INTERFACE ITF_Buffer2_4

METHOD Aborted : BOOL
VAR_INPUT
END_VAR
END_METHOD

METHOD Aborting : BOOL
VAR_INPUT
END_VAR
END_METHOD

METHOD Clearing : BOOL
VAR_INPUT
END_VAR
END_METHOD

METHOD Execute : BOOL
VAR_INPUT
END_VAR
END_METHOD

METHOD Held : BOOL
VAR_INPUT
END_VAR
END_METHOD

METHOD Holding : BOOL
VAR_INPUT
END_VAR
END_METHOD

METHOD Idle : BOOL
VAR_INPUT
END_VAR
END_METHOD

METHOD Resetting : BOOL
VAR_INPUT
END_VAR
END_METHOD

METHOD Starting : BOOL
VAR_INPUT
END_VAR
END_METHOD

METHOD Stopped : BOOL
VAR_INPUT
END_VAR
END_METHOD

METHOD Stopping : BOOL
VAR_INPUT
END_VAR
END_METHOD

METHOD Suspended : BOOL
VAR_INPUT
END_VAR
END_METHOD

METHOD Suspending : BOOL
VAR_INPUT
END_VAR
END_METHOD

METHOD Unholding : BOOL
VAR_INPUT
END_VAR
END_METHOD

METHOD Unsuspending : BOOL
VAR_INPUT
END_VAR
END_METHOD

END_INTERFACE

(* stored: Version 1.1.0.1
   Itf ITF_Buffer2_4: Id {b287fb4f-1856-4601-beeb-92f66b9fe064}
   Folder Methods: Id {e87007a4-9015-4af8-9b6c-24c986ad8a52}
   Method Aborted: Id {23f30cc0-5225-4a77-ba8d-ab499bbc1a2a}
   Method Aborting: Id {39ac2970-0f2e-4beb-9e13-3f810caf740b}
   Method Clearing: Id {a14ccadc-97d7-4a07-8c73-39905745d9b0}
   Method Execute: Id {1ceb5459-e1ba-49c9-b800-d68fb4dc205a}
   Method Held: Id {fb6cae87-1391-46f9-930d-e4581e1b4bc4}
   Method Holding: Id {5219f426-63fa-49ce-9216-8264765adf30}
   Method Idle: Id {4f6d92b3-e523-4cc6-8396-0ba2c86a8cff}
   Method Resetting: Id {df32f635-75c3-4076-842c-d7e80f85be61}
   Method Starting: Id {6817a570-5ca6-4f55-a121-e387572f434e}
   Method Stopped: Id {232b9b6b-9f09-4086-8b7b-bf7cb90e0b93}
   Method Stopping: Id {20ba74bf-8da2-47eb-84e9-a2625a31e303}
   Method Suspended: Id {ac324cdd-6861-4f12-b6e8-847cf360fe5b}
   Method Suspending: Id {3f96b2d4-44c9-45ec-a31f-ad6577ca7690}
   Method Unholding: Id {e59049e1-536e-4a9c-b3c3-d015b3de706d}
   Method Unsuspending: Id {9406f3f1-76a1-4fff-a5e0-19a8f19015d8} *)
